{attribute 'qualified_only'}
{attribute 'strict'}
TYPE E_Parameters :
(
	isLoggerEnabled 				:= 1,
	cylinderTimeout					:= 2,
//	airPressureMin					:= 3,
//	airPressureMax					:= 4,
	numberOfRetries					:= 5
	
);
END_TYPE

(* stored: Version 1.1.0.1, ProductVersion 3.1.4024.12
   DUT E_Parameters: Id {7f6c40a4-0a35-0199-37b8-9aea5080de17} *)
